# EPICS substitutions: db/Beckhoff_1XXX/ecmcEP1258.substitutions
# binary inputs
file "ecmc_binaryInput-chX.template"{
  pattern {CH_ID}
          {01   }
          {02   }
          {03   }
          {04   }
          {05   }
          {06   }
          {07   }
          {08   }
}

# timestamp, only channel 1 and 2 have this feature
file "ecmc_timestamp_64-chX.template"{
  pattern {CH_ID, KEY,          suffix,  sourceName                }
          {01,    "BI",  "-TimeRise",    "timestampLatchPositive"  }
          {01,    "BI",  "-TimeFall",    "timestampLatchNegative"  }
          {02,    "BI",  "-TimeRise",    "timestampLatchPositive"  }
          {02,    "BI",  "-TimeFall",    "timestampLatchNegative"  }
}

# channel status
file "ecmc_status-chX.template"{
  pattern {CH_ID, KEY}
          {01,    BI }
          {02,    BI }
}
